(* PLC project Vn_ld_parallel3, Beckhoff Automation GmbH TwinCAT PLC Control 3.5.13.21 *)
(* stored: creationDateTime 1970-01-01T00:00:00 *)

PROGRAM Vn_ld_parallel3

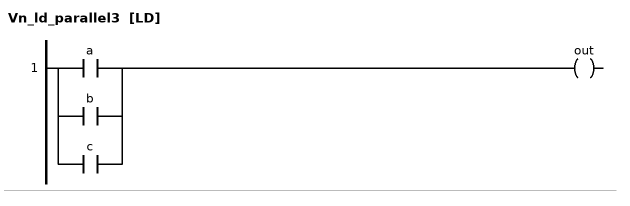
(* LD diagram, written out as Structured Text *)
out := a OR b OR c;
END_PROGRAM
